// Mitsubishi GX Works2 project: 261012_기초회로_비상정지회로   PLC: Q03UDV

PROGRAM MAIN
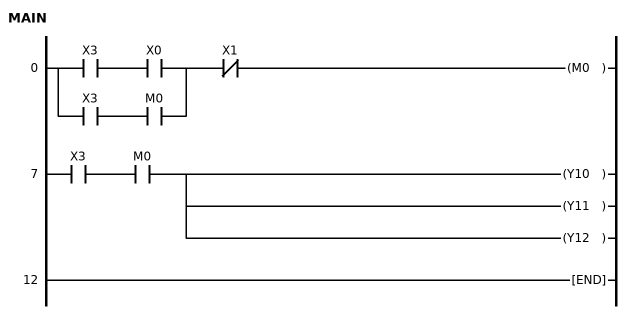
0     LD      X3
      AND     X0
      LD      X3
      AND     M0
      ORB
      ANI     X1
      OUT     M0
7     LD      X3
      AND     M0
      OUT     Y10
      OUT     Y11
      OUT     Y12
12    END
END_PROGRAM
